Staubli VAL3: setnullmode.pgx

public program setnullmode()
  local num l_i
begin
  $jogMode(0)
   for l_i = 0 to size(sShowType)-1
    sShowType[l_i]=sCartisiam[l_i]
  endFor
end
